// TIA Portal V20 export
// export: Created 2026-10-12T16:46:21.3656708Z, ExportSetting WithDefaults, DisplayName Totally Integrated Automation Portal, DisplayVersion V20 Update 6, DisplayName TIA Portal Openness, DisplayVersion V20 Update 6, DisplayName TIA Portal Version Control Interface, DisplayVersion V20 Update 6, DisplayName SINAMICS Startdrive Advanced, DisplayVersion V20 SP1 Update 2, DisplayName SINAMICS Startdrive G110M, G120, G120C, G120D, G120P, G115D, DisplayVersion V20 SP1 Update 2, DisplayName SINAMICS Startdrive G130, G150, S120, S150, SINAMICS MV, G220, S200, S210, DisplayVersion V20 SP1 Update 2, DisplayName STEP 7 Professional, DisplayVersion V20 Update 6, DisplayName STEP 7 Safety, DisplayVersion V20 Update 2, DisplayName WinCC Basic/Comfort/Advanced, DisplayVersion V20 Update 6, DisplayName WinCC Professional, DisplayVersion V20 Update 6, DisplayName WinCC Unified, DisplayVersion V20 Update 6
DATA_BLOCK "DB_HMI"   // DB4
{ S7_Optimized_Access := 'TRUE' }
VERSION : 0.1
// stored: AutoNumber true, DBAccessibleFromOPCUA true, DBAccessibleFromWebserver true, IsOnlyStoredInLoadMemory false, IsRetainMemResEnabled false, IsWriteProtectedInAS false, MemoryReserve 100
   VAR
      Benutzerverwaltung_User_Daten { S7_SetPoint := 'True'} : "UDT_Benutzer";
      Benutzerverwaltung_User_create { S7_SetPoint := 'True'} : Bool;
      Benutzerverwaltung_User_update : Bool;
      Benutzerverwaltung_User_delete : Bool;
      Benutzerverwaltung_Freigaben_Prozessgruppen_User_change : Bool;
      Benutzerverwaltung_Status : Int;
      Benutzerverwaltung_Freigabe_Prozessgruppen_User_ID_ausgewählt : Int;
      Benutzerverwaltung_Freigabe_Prozessgruppen_Prozessgruppen : Array[1.."c_Prozessgruppen"] of Bool;
      Benutzerverwaltung_Login_Name : String;
      Benutzerverwaltung_Login_Passwort : String;
      Benutzerverwaltung_Login_Loginbutton : Bool;
      Benutzerverwaltung_Login_Logoutbutton : Bool;
      Benutzerverwaltung_Login_Login_Ok : Bool;
      Prozessparameter_Status : Int;
      Prozessparameter_Prozessgruppen_save : Bool;
      Prozessparameter_Prozessgruppen_Prozessgruppe : "UDT_Prozessgruppen";
      Prozessparameter_Artikel_add { S7_SetPoint := 'True'} : "UDT_Artikel";
      Prozessparameter_Artikel_save { S7_SetPoint := 'True'} : Bool;
      Prozessparameter_Artikel_delete : Bool;
      Prozessparameter_Artikel_assign : Bool;
      Prozessparameter_Artikel_remove : Bool;
      "Prozessparameter_Prozessgruppe_ID_assign/remove" : Int;
      "Prozessparameter_Artikel_ID_assign/remove" : Int;
      Angewähltes_Bad : USInt;
      Handbetrieb { S7_SetPoint := 'True'} : "UDT_Handbetrieb";
   END_VAR
BEGIN
END_DATA_BLOCK
